FUNCTION_BLOCK FB_Blinker
VAR_INPUT
	bStart: BOOL;
	tSignalTimerOn: TIME;
	tSignalTimerOff: TIME;
END_VAR
VAR_OUTPUT
	bOut: BOOL;
END_VAR
VAR
	fbTimerA: TON;
	fbTimerB: TON;
END_VAR

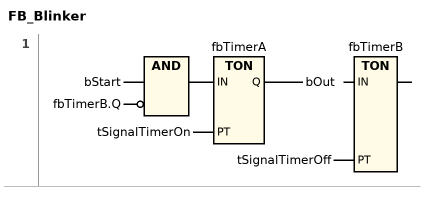
// NETWORK 1
fbTimerA(IN := bStart AND NOT fbTimerB.Q, PT := tSignalTimerOn); // TON
bOut := fbTimerA.Q;
fbTimerB(IN := fbTimerA.Q, PT := tSignalTimerOff); // TON

END_FUNCTION_BLOCK

(* stored: Version 1.1.0.1, ProductVersion 3.1.4024.16
   POU FB_Blinker: Id {c4623b14-e343-46ac-bdaa-ca112f838f7e}, SpecialFunc None *)
